// Mitsubishi GX Works2 project: 시험1_테스트동작   PLC: FX3U/FX3UC

PROGRAM MAIN
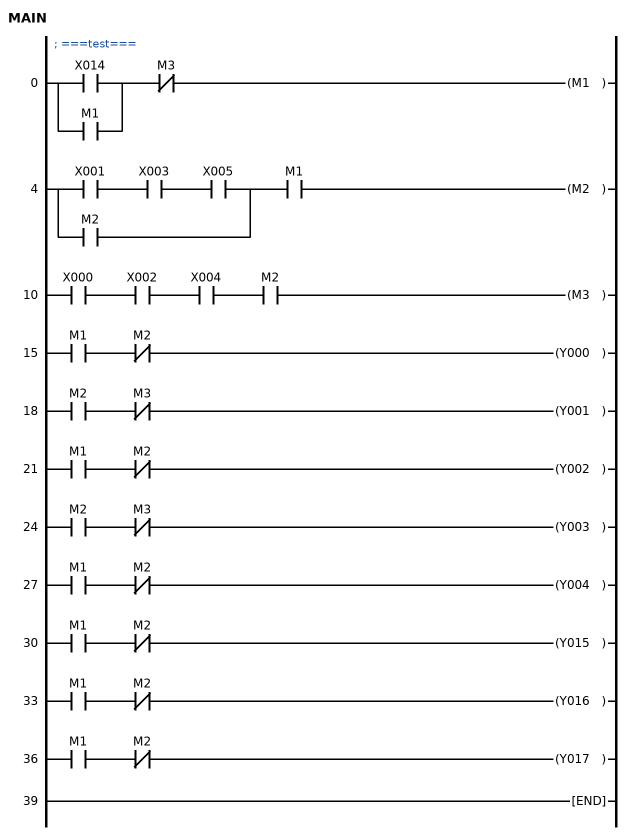
; ===test===
0     LD      X014
      OR      M1
      ANI     M3
      OUT     M1
4     LD      X001
      AND     X003
      AND     X005
      OR      M2
      AND     M1
      OUT     M2
10    LD      X000
      AND     X002
      AND     X004
      AND     M2
      OUT     M3
15    LD      M1
      ANI     M2
      OUT     Y000
18    LD      M2
      ANI     M3
      OUT     Y001
21    LD      M1
      ANI     M2
      OUT     Y002
24    LD      M2
      ANI     M3
      OUT     Y003
27    LD      M1
      ANI     M2
      OUT     Y004
30    LD      M1
      ANI     M2
      OUT     Y015
33    LD      M1
      ANI     M2
      OUT     Y016
36    LD      M1
      ANI     M2
      OUT     Y017
39    END
END_PROGRAM
